(* IEC 61131-3 sources: volt/packages/volt-lsp-iec/test-corpus/awa-palletizer/Device/Plc Logic/Application/Library Manager/L_IE1P_ApplicationErrorsTypes, 22 files *)

(* ---- L_IE1P_ERROR.dut ---- *)
TYPE L_IE1P_ERROR :
(
	NOERROR := 0,
	MODULOAXISISREQUIRED := 17000,
	STARTPOSOUTOFCYCLELENGTH := 17003,
	CYCLELENGHTSHAVETOBEEQUAL := 17004,
	INVALIDDIRECTION := 17005,
	MARKSTACKLIMITREACHED := 17006,
	MAXMISSEDMARKS := 17007,
	INVALIDFOLLOWLINEACCVEL := 17008,
	INVALIDJOGGINGACCVEL := 17009,
	INVALIDSTOPDEC := 17010,
	INVALIDDIAMETER := 17011,
	TORQUEFOLLOWERNOTREADYFORMOTION := 17012,
	SPEEDFOLLOWERNOTREADYFORMOTION := 17013,
	INVALIDINVERTER := 17014,
	SDO_ACCESSFAILEDTOMOTORPARAMETERS := 17015,
	MISSEDMAPPINGPARAMETERLOWERSPEEDLIMIT := 17016,
	MISSEDMAPPINGPARAMETERUPPERSPEEDLIMIT := 17017,
	MISSEDMAPPINGPARAMETERTORQUEOFFSET := 17018,
	DANCERPOSOUTOFRANGE := 17019,
	INVALIDLIMITDANCERPOS := 17020,
	INVALIDCLUTCHPARAMETERS := 17021,
	WASNOTCALLEDDURINGMOTION := 17022,
	INVALIDNUMBEROFCAMPOINTS := 17030,
	INVALIDPATHPAR := 17032,
	INVALIDBLENDINGRADIUS := 17033,
	PATHNOTSUPPORTED := 17034,
	X_PATHLIMITPOSITIVEEXCEEDED := 17035,
	X_PATHLIMITNEGATIVEEXCEEDED := 17036,
	Y_PATHLIMITPOSITIVEEXCEEDED := 17037,
	Y_PATHLIMITNEGATIVEEXCEEDED := 17038,
	Z_PATHLIMITPOSITIVEEXCEEDED := 17039,
	Z_PATHLIMITNEGATIVEEXCEEDED := 17040,
	C_PATHLIMITPOSITIVEEXCEEDED := 17041,
	C_PATHLIMITNEGATIVEEXCEEDED := 17042,
	INVALIDPATHDATA := 17043,
	INVALIDTARGETPLC := 17047,
	MINLIMITVELGTPROFILEVEL := 17048,
	MINLIMITACCGTPROFILEACC := 17049,
	MINLIMITDECGTPROFILEDEC := 17050,
	MASTERISMOVING := 17100,
	INVALIDPODUCTLENGTH := 17101,
	TPSENSORNOTTEACHED := 17102,
	SLAVERECEIVEDGAPS := 17103,
	MASTERRECEIVEDGAPS := 17104,
	INTERNALERROR := 17105,
	INVALIDPARAMETERCUTTINGANGLE := 17106,
	INVALIDCUTTINGPARAMETERS := 17107,
	INVALIDCUTTINGLENGTH := 17108,
	SLAVENOTINPARKPOS := 17109,
	MASTERISREVERSING := 17110,
	INTINVALIDSELECTCAM := 17111,
	SELECTEDAXISISNOTSUPPORTED := 17112,
	AXISISNOTSUPPORTED := 17113,
	INVALIDPROFILE := 17114,
	AXISENABLEDISREQUIRED := 17115,
	CORRLIMITOUTOFCYCLELENGTH := 17116,
	CORRECTIONGREATERCORRWINDOW := 17117,
	INVALIDCNCPROGRAM := 17118,
	SAFEDISTVIOLATION := 17119,
	SAFEDISTINSUFFICIENTFORSTOP := 17120,
	INVALIDGCODELINE := 17121,
	COORDSYSTEMACSNOTSUPPORTED := 17122,
	DANCERLIMITSNOTTEACHED := 17123,
	NOTREADYFORADDPROFILE := 17124,
	SLAVEPOSUPPERLIMIT := 17125,
	SLAVEPOSLOWERLIMIT := 17126,
	TARGETPOSUPPERLIMIT := 17127,
	INVALIDMARKPOSITION := 17128,
	INVALIDPOSITIONINGMODE := 17129,
	TEMPSENSORFAILURE := 17130,
	MAXCRITICALTEMPREACHED := 17131,
	INVALIDTEMPCONTROLPARAM := 17132,
	IDENTIFICATIONFAILED := 17133,
	PWMTASKCYCLEMISMATCH := 17134,
	CONCURRENTREQUESTTEMPCONTROL := 17135,
	TMNOTCALLEDINCYCLICTASK := 17136,
	TMDATABUSDISCONNECTED := 17137,
	INVALIDTMDATABUS := 17138,
	TMDATABUSCONFIGCHANGED := 17139,
	TMNOTCALLEDINMOTIONTASK := 17140,
	SLAVETMSTATESERVICE := 17141,
	COLLISIONDETECTIONDISABLED := 17142,
	COLLISIONDETECTED := 17143,
	INVALIDTMDATABUSORDER := 17144,
	CHANGEOFCONVEYORAXESNOTALLOWED := 17145,
	INVALIDSETTARGET := 17146,
	LOWERLIMITEXCEEDSUPPERLIMIT := 17147,
	SETTARGETSTACKLIMITREACHED := 17148,
	WORKPIECESTACKLIMITREACHED := 17149,
	INVALIDTRAVERSINGPROFILEPARAMETER := 17150,
	INVALIDTRAVERSINGCOILPARAMETER := 17151,
	TRAVERSINGANGULARSHIFTLIMITREACHED := 17152,
	AXESGROUPALREADYINUSE := 17153,
	UNDERVOLTAGEDCLINK := 17154,
	COUPLINGMODEREQUIRESMODULOAXIS := 17155,
	DUPLICATEDTM_ADDRESS := 17156,
	XAXISTMERROR := 17157,
	YAXISTMERROR := 17158,
	APAXISTMERROR := 17159,
	SLAVEXAXISTMERROR := 17160,
	SLAVEYAXISTMERROR := 17161,
	INVALIDMOVEPPACTIVE := 17162,
	INVALIDCONVEYORBELTPAR := 17163,
	IDENTIFICATIONDIAMETERFAILED := 17164,
	ACTDANCERPOSGTMAXDANCERPOS := 17165,
	INVALIDIDENTMAXDANCERPOS := 17166,
	INVALIDDANCERMATERIALLENGTH := 17167,
	LOADDIAMETERNOTALLOWED := 17168,
	INVALIDMASTERAXISREF := 17169,
	SYNCMODEVELACCREQUIRED := 17170,
	TEMPMAXCRITICALEXCEEDED := 17171,
	INVALIDTEMPCTRLPARAM := 17172,
	INVALIDSYNCSLAVEDIRECTION := 17173,
	MARKCORRECTIONINNEXTCYCLE := 17174,
	BASEVELOCITYNOTSUPPORTED := 17175,
	MOVEMENTBLOCKEDBYTRAINAHEAD := 17176,
	MARKDISTANCEGTZEROREQUIRED := 17177,
	INVALIDVIRTMASTERSETVELZERO := 17178,
	HOMINGBLOCKEDBYACTIVEFUNCTION := 17179,
	CONCURRENTMOTIONCMDDURINGHOMING := 17180,
	INVALIDCYCLELENGTHETCONBOARD := 17181,
	INVALIDMASTERVALUESOURCE := 17182,
	ETCONBOARDNOTOPERATIONAL := 17183,
	TRAVERSINGRANGEMASTERNOTEQUALVIRTMASTER := 17184,
	CYCLELENGTHMASTERNOTEQUALVIRTMASTER := 17185,
	MISSEDMAPPINGPARAMETERTPTIMESTAMP := 17186,
	TOLERANCEALLOWEDDIRECTIONEXCEEDED := 17187,
	TPRECPOSITIONNOTSUPPORTED := 17188,
	INVALIDHYSTERESISWIDTH := 17189,
	ALLOWEDDIRECTIONVIOLATEDBYBASEVELOCITY := 17190,
	VELOUTOFTOLERANCEINVERTGEARFACTOR := 17191,
	INVALIDPARAMETERCOMBINATIONACDRIVEPROFILE := 17192,
	MINVELLIMITGTMAXVELLIMIT := 17193,
	SETVALUEMODENOTSUPPORTED := 17194,
	LINEVELDIAMCALCREQUIRED := 17195,
	INVALIDSTOPMODE := 17196,
	INVALIDDIRECTIONFORTARGETMATERIALCOUNTER := 17197,
	MAXMISSEDMARKSTOOL := 17198,
	MODECHANGEBLOCKEDBYSYNCIN := 17199,
	CONCURRENTMOTIONCMDDURINGSERVICE := 17200,
	STOPPOSITIONEXCEEDED := 17201,
	NOTREADYFORCOORDINATEDMOTION := 17202,
	INVALIDMARKWINDOWMASTERVALUECORR := 17203,
	INVALIDMARKWINDOWTOOLCORR := 17204,
	FUNCTIONBLOCKEDBYTRAVERSING := 17205,
	MASTERCYCLELENGTHCHANGED := 17206,
	TRIMMINGONLYDURINGSYNCHRONISED := 17207,
	LOWERTURNPOSGTUPPERTURNPOS := 17208,
	MASTERNOTCONNECTED := 17209,
	CANNOTCATCHUP := 17210,
	MISSINGMMADDRESS := 17901,
	NUMOFMMEXCEEDED := 17902,
	DUPLICATEDROOTMM := 17903,
	SLAVEMMNOTFOUND := 17904,
	ZPOSMAXEXCEEDED := 17905,
	MISSINGMODULEREFERENCE := 17906,
	ERRORLISTOVERFLOW := 17907,
	ACDOWNSTRUCTINVALID := 17908,
	ACDSLAVESTRUCTINVALID := 17909,
	ACDSIZEOVERFLOW := 17910,
	COMPIDOUTOFRANGE := 17911,
	TOOMANYLEVELS := 17912,
	MMDSTRUCTINVALID := 17913,
	NOPOOLRESOURCEAVAILABLE := 17914,
	NORESOURCEMOVELINABS := 17915,
	NORESOURCEMOVELINREL := 17916,
	NORESOURCEMOVEDIRABS := 17917,
	NORESOURCEMOVEDIRREL := 17918,
	NORESOURCEPNP := 17919,
	NOCOMMANDRECEIVERAVAILABLE := 17920,
	COMMANDRECEIVERNOTENABLED := 17921,
	INTERNALCONTROLACTIVE := 17922,
	INTERNALCONTROLENABLED := 17923,
	INTERNALCONTROLDISABLED := 17924,
	MMCOUPLINGDISABLED := 17925,
	MMCOUPLINGENABLED := 17926,
	MODECHANGEREQUESTED := 17927,
	MODENUMBEROUTSIDERANGE := 18001,
	MODENUMBERNOTUSEDINCONFIG := 18002,
	MODECHANGENOTALLOWEDINCURRENTMODE := 18003,
	MODECHANGENOTALLOWEDINNEXTMODE := 18004,
	LI_MODENUMBEROUTSIDERANGE := 18005,
	LI_MODENUMBERNOTUSEDINCONFIG := 18006,
	LI_MODECHANGENOTALLOWEDREMOTE := 18007,
	LI_MODECHANGENOTALLOWEDINCURRENTMODE := 18008,
	LI_MODECHANGENOTALLOWEDINNEXTMODE := 18009,
	MORETHANONECOMMANDACTIVE := 18010,
	CONCURRENTCOMMAND := 18011,
	COMMANDNOTALLOWEDINCURRENTSTATE := 18012,
	LI_COMMANDSONLYINMODEPRODUCTION := 18013,
	LI_COMMANDNOTALLOWEDINREMOTE := 18014,
	LI_COMMANDNOTALLOWEDINCURRENTSTATE := 18015,
	CONCURRENTTOOLCMD := 18016,
	DELAYTIMEINVALID_PT1FILTER := 19000,
	MODEINVALID_CURVE := 19002,
	MODEINVALID_COMPARE := 19003,
	MODEINVALID_CONVAXISV := 19005,
	DELAYTIMEINVALID_PROCESSCONTROLLER := 19006,
	RATETIMEINVALID_PROCESSCONTROLLER := 19007,
	RESETTIMEINVALID_PROCESSCONTROLLER := 19008,
	MODEINVALID_DELAY := 19024,
	ABORTEDBYSTARTIDENT_FRICTCOMP := 19030,
	ABORTEDBYFOLLOWERDISABLED_FRICTCOMP := 19031,
	MAXSPEEDNOTREACHED_FRICTCOMP := 19032,
	ACCTOOBIG_FRICTCOMP := 19033,
	DMINBIGGERDMAX_CALCDIAMETER := 19034,
	MAXSPEEDORMAXTORQUE_IDENTMINERTIA := 19048,
	ABORTEDBYSTARTIDENT_IDENTMINERTIA := 19049,
	ABORTEDBYFOLLOWERDISABLED_IDENTMINERTIA := 19050,
	ABORTEDBYFOLLOWERENABLED_IDENTMINERTIA := 19051,
	NMAXNOTREACHED_IDENTMINERTIA := 19052,
	MNOTREACHED_IDENTMINERTIA := 19053,
	MAXNROFTPEXCEEDED_MARKREGISTER := 19503,
	IDENTMODENOTSUPPORTED := 19801,
	MOTORRATEDSPEEDZERO := 19803,
	INERTIAMOTORZERO := 19804,
	STARTMODEINVALID := 19806,
	INVALIDEIGENFREQUENCY := 19807,
	INVALIDAMPLITUDERATIO := 19808,
	INVALIDOSCCOMPMODE := 19809,
	CHANGEOFOSCCOMPMODELOCKED := 19810,
	INVALIDDEFAULTCONTROLMODE := 19812,
	INVALIDMOTORCONTROLMODE := 19813,
	VIRTUALMODENOTALLOWED := 19814,
	POSITIONWINDOWNEGOUTSIDESWLIMITS := 19817,
	POSITIONWINDOWPOSOUTSIDESWLIMITS := 19818,
	ACTPOSITIONOUTSIDEWINDOW := 19819,
	PROFILEEXCEEDSPOSITIONWINDOW := 19820,
	ACTVELOCITYEXCEEDSTOLERANCE := 19822,
	ACTTORQUEEXCEEDSTOLERANCE := 19823,
	POSITIONWINDOWNEGVIOLATION := 19825,
	POSITIONWINDOWPOSVIOLATION := 19826,
	AXISINSTABILITYDUETOSTARTCTRLPARAM := 19827,
	INPOSITIONTIMEOUT := 19828,
	RESTOREDATANOTAVAILABLE := 19829,
	POSITIONWINDOWREQUIRESLIMITEDAXIS := 19830,
	MISSEDMAPPINGPARAMETERVELOCITYERROR := 19831,
	INSTABILITYDUETOTUNESTRATEGY := 19832,
	ARRAYBOUNDSNOTEQUALMODULOCYCLE := 19833,
	PERIODICCORRECTIONVALUESREQUIRED := 19834,
	INVALIDBACKLASHCOMPMODE := 19835,
	INVALIDBACKLASHWIDTH := 19836,
	INVALIDCOMPTIME := 19837,
	BACKLASHWIDTHGTCYCLELENGTH := 19838,
	SDO_OTHERERROR := 20001,
	SDO_INVALIDINDEX := 20002,
	SDO_INVALIDOFFSET := 20003,
	SDO_INVALIDSIZE := 20004,
	SDO_INVALIDDATA := 20005,
	SDO_NOTREADY := 20006,
	SDO_BUSY := 20007,
	SDO_NOMEMORY := 20008,
	SDO_INVALIDPARM := 20009,
	SDO_INVALIDSTATE := 20010,
	SDO_TIMEOUT := 20011,
	SDO_INVALID_SLAVE_STATE := 20012,
	SDO_LINK_DISCONNECTED := 20013,
	SDO_ALL_CANNELS_BUSY := 20015,
	SDO_ABORTCODE_TOGGLE := 20020,
	SDO_ABORTCODE_TIMEOUT := 20021,
	SDO_ABORTCODE_CCS_SCS := 20022,
	SDO_ABORTCODE_BLK_SIZE := 20023,
	SDO_ABORTCODE_SEQNO := 20024,
	SDO_ABORTCODE_CRC := 20025,
	SDO_ABORTCODE_MEMORY := 20026,
	SDO_ABORTCODE_ACCESS := 20027,
	SDO_ABORTCODE_WRITEONLY := 20028,
	SDO_ABORTCODE_READONLY := 20029,
	SDO_ABORTCODE_INDEX := 20030,
	SDO_ABORTCODE_PDO_MAP := 20031,
	SDO_ABORTCODE_PDO_LEN := 20032,
	SDO_ABORTCODE_P_INCOMP := 20033,
	SDO_ABORTCODE_I_INCOMP := 20034,
	SDO_ABORTCODE_HARDWARE := 20035,
	SDO_ABORTCODE_DATA_SIZE := 20036,
	SDO_ABORTCODE_DATA_SIZE1 := 20037,
	SDO_ABORTCODE_DATA_SIZE2 := 20038,
	SDO_ABORTCODE_OFFSET := 20039,
	SDO_ABORTCODE_DATA_RANGE := 20040,
	SDO_ABORTCODE_DATA_RANGE1 := 20041,
	SDO_ABORTCODE_DATA_RANGE2 := 20042,
	SDO_ABORTCODE_MINMAX := 20043,
	SDO_ABORTCODE_GENERAL := 20044,
	SDO_ABORTCODE_TRANSFER := 20045,
	SDO_ABORTCODE_TRANSFER1 := 20046,
	SDO_ABORTCODE_TRANSFER2 := 20047,
	SDO_ABORTCODE_DICTIONARY := 20048,
	SDO_ABORTCODE_UNKNOWN := 20049,
	NOAXISREF := 20301,
	NOPARAMETER := 20302,
	NOVALIDPARAM := 20303,
	NOVALIDAXISSTATE := 20304,
	NOBOOLPARAM := 20305,
	SWLIMITPOS := 20306,
	SWLIMITNEG := 20307,
	NOVALID_MC_SOURCE := 20308,
	NOSETVALUESAVAILABLE := 20309,
	POWERFAILDURINGOPERATION := 20310,
	NOTREADYFORMOTION := 20311,
	POSSWLIMITREACHED := 20312,
	NEGSWLIMITREACHED := 20313,
	NOVALIDTPSOURCE := 20314,
	NOVALIDTPNUMBER := 20315,
	TPALREADYACTIVE := 20316,
	NOTTPSUPPORTED := 20317,
	NOTPACTIVE := 20318,
	NOEXTPINPUT := 20319,
	NOVALIDACCELERATION := 20320,
	NOVALIDDECELERATION := 20321,
	NOVALIDVELOCITY := 20322,
	ARITHMETICERROR := 20323,
	NOTAPPLICABLE := 20324,
	VELOCITYLIMITED := 20325,
	ACCELERATIONLIMITED := 20326,
	JERKLIMITED := 20327,
	TARGETOUTSIDESWLIMIT := 20328,
	JERKLIMITATIONDEACTIVATEDDUETOARITHMETICERROR := 20329,
	NOVALIDACCELERATION_MOVEABSOLUTE := 20330,
	NOVALIDDECELERATION_MOVEABSOLUTE := 20331,
	NOVALIDVELOCITY_MOVEABSOLUTE := 20332,
	ARITHMETICERROR_MOVEABSOLUTE := 20333,
	NOTAPPLICABLE_MOVEABSOLUTE := 20334,
	VELOCITYLIMITED_MOVEABSOLUTE := 20335,
	ACCELERATIONLIMITED_MOVEABSOLUTE := 20336,
	JERKLIMITED_MOVEABSOLUTE := 20337,
	TARGETOUTSIDESWLIMIT_MOVEABSOLUTE := 20338,
	NOVALIDACCELERATION_MOVEADDITIVE := 20340,
	NOVALIDDECELERATION_MOVEADDITIVE := 20341,
	NOVALIDVELOCITY_MOVEADDITIVE := 20342,
	ARITHMETICERROR_MOVEADDITIVE := 20343,
	NOTAPPLICABLE_MOVEADDITIVE := 20344,
	VELOCITYLIMITED_MOVEADDITIVE := 20345,
	ACCELERATIONLIMITED_MOVEADDITIVE := 20346,
	JERKLIMITED_MOVEADDITIVE := 20347,
	TARGETOUTSIDESWLIMIT_MOVEADDITIVE := 20348,
	NOVALIDACCELERATION_MOVECONTAB := 20350,
	NOVALIDDECELERATION_MOVECONTAB := 20351,
	NOVALIDVELOCITY_MOVECONTAB := 20352,
	ARITHMETICERROR_MOVECONTAB := 20353,
	NOTAPPLICABLE_MOVECONTAB := 20354,
	VELOCITYLIMITED_MOVECONTAB := 20355,
	ACCELERATIONLIMITED_MOVECONTAB := 20356,
	JERKLIMITED_MOVECONTAB := 20357,
	TARGETOUTSIDESWLIMIT_MOVECONTAB := 20358,
	NOVALIDACCELERATION_MOVECONTREL := 20360,
	NOVALIDDECELERATION_MOVECONTREL := 20361,
	NOVALIDVELOCITY_MOVECONTREL := 20362,
	ARITHMETICERROR_MOVECONTREL := 20363,
	NOTAPPLICABLE_MOVECONTREL := 20364,
	VELOCITYLIMITED_MOVECONTREL := 20365,
	ACCELERATIONLIMITED_MOVECONTREL := 20366,
	JERKLIMITED_MOVECONTREL := 20367,
	TARGETOUTSIDESWLIMIT_MOVECONTREL := 20368,
	NOVALIDACCELERATION_MOVERELATIVE := 20370,
	NOVALIDDECELERATION_MOVERELATIVE := 20371,
	NOVALIDVELOCITY_MOVERELATIVE := 20372,
	ARITHMETICERROR_MOVERELATIVE := 20373,
	NOTAPPLICABLE_MOVERELATIVE := 20374,
	VELOCITYLIMITED_MOVERELATIVE := 20375,
	ACCELERATIONLIMITED_MOVERELATIVE := 20376,
	JERKLIMITED_MOVERELATIVE := 20377,
	TARGETOUTSIDESWLIMIT_MOVERELATIVE := 20378,
	NOVALIDACCELERATION_MOVESUPERIMP := 20380,
	NOVALIDDECELERATION_MOVESUPERIMP := 20381,
	NOVALIDVELOCITY_MOVESUPERIMP := 20382,
	ARITHMETICERROR_MOVESUPERIMP := 20383,
	NOTAPPLICABLE_MOVESUPERIMP := 20384,
	VELOCITYLIMITED_MOVESUPERIMP := 20385,
	ACCELERATIONLIMITED_MOVESUPERIMP := 20386,
	JERKLIMITED_MOVESUPERIMP := 20387,
	TARGETOUTSIDESWLIMIT_MOVESUPERIMP := 20388,
	NOVALIDACCELERATION_MOVEVELOCITY := 20390,
	NOVALIDDECELERATION_MOVEVELOCITY := 20391,
	NOVALIDVELOCITY_MOVEVELOCITY := 20392,
	ARITHMETICERROR_MOVEVELOCITY := 20393,
	NOTAPPLICABLE_MOVEVELOCITY := 20394,
	VELOCITYLIMITED_MOVEVELOCITY := 20395,
	ACCELERATIONLIMITED_MOVEVELOCITY := 20396,
	JERKLIMITED_MOVEVELOCITY := 20397,
	TARGETOUTSIDESWLIMIT_MOVEVELOCITY := 20398,
	NOVALIDDECELERATION_HALT := 20401,
	ARITHMETICERROR_HALT := 20403,
	ACCELERATIONLIMITED_HALT := 20406,
	JERKLIMITED_HALT := 20407,
	NOVALIDDECELERATION_STOP := 20411,
	ARITHMETICERROR_STOP := 20413,
	ACCELERATIONLIMITED_STOP := 20416,
	JERKLIMITED_STOP := 20417,
	NOVALIDDIRECTION := 20430,
	NOVALIDBUFFERMODE := 20431,
	DIRECTIONDISABLED := 20432,
	BLOCKEDBYAXISSTATE := 20433,
	NOVALIDOVERRIDE := 20434,
	CONCURRENT_MC_POWER := 20435,
	CONCURRENT_SETQUICKSTOP := 20436,
	FDBABSPOSNOTAVAILABLE := 20498,
	DRIVE_PDO_INTERFACE_DISABLED := 20499,
	HWLIMITPOS := 20500,
	HWLIMITNEG := 20501,
	FOLLOWINGERROR1 := 20502,
	FOLLOWINGERROR2 := 20503,
	COMMUNICATIONFAIL := 20504,
	AXISINITFAIL := 20505,
	COMMTIMOUT := 20506,
	MASTERRESTARTFAIL := 20507,
	NOTREADYFORREINIT := 20508,
	ERRORDURINGINIT := 20509,
	SWITCHONNOTPOSSIBLE := 20510,
	DRIVEERROR := 20511,
	HOME_NOAUXPARAMETERS := 20512,
	HOME_MODENOTSUPPORTEDBYAXIS := 20513,
	HOME_MODEUNKNOWN := 20514,
	HOME_NOAUXTRIGGERINPUT := 20515,
	HOME_UNKNOWNTPCONFIG := 20516,
	HOME_WRITEHOMEPARAMETER := 20518,
	HOME_ERRORWHILEHOMING := 20519,
	HOME_ARITHMETICERROR := 20520,
	HOME_TORQUELIMNOTMAPPED := 20521,
	HOME_INVALIDVELACC := 20522,
	HOMETPEDGESETTINGNOTSUPPORTED := 20523,
	RESETDRIVEERRORFAILED := 20525,
	APPLICATIONERROR := 20526,
	APPLICATIONWARNING := 20527,
	BRAKE_POSITIONDRIFT := 20529,
	BRAKE_INVALIDMODE := 20530,
	BRAKE_TIMEOUTPRECONTROL := 20531,
	BRAKE_INVALIDBRAKESTATE := 20532,
	FAST_IO_OUT_WRONGOUTPUTSEL := 20533,
	FAST_IO_OUT_NOFREEENCODERAXIS := 20534,
	FAST_IO_OUT_FREEENCODERAXISWRONGPARAMETER := 20535,
	FAST_IO_OUT_MAPPINGFAULT := 20536,
	FAST_IO_OUT_FIFOOVERFLOW := 20537,
	TP_SELECT := 20538,
	TP_MODE := 20539,
	TP_ONLYPOSEDGE := 20540,
	TP_EDGENOTAVAILABLE := 20541,
	TP_CHANNELNOTFREE := 20542,
	TP_MAPPINGFAULT := 20543,
	TP_INTERNALCHANNELNOTFREE := 20544,
	TP_TIMEOUT := 20545,
	TP_COMMUNICATIONERROR := 20546,
	TP_SIGNAL := 20547,
	TP_NOFREEENCODERAXIS := 20548,
	TP_PARAMETERRISINGEDGEWRONGVALUE := 20550,
	TP_PARAMETERFALLINGRISINGEDGEWRONGVALUE := 20551,
	TP_INTERNALERROR := 20552,
	SETVALUESGTMAXAPPVALUES := 20600,
	SETVALUESINCONSISTENT := 20601,
	POSDIFFGTHALFCYCLELENGTH := 20602,
	INVALIDTASKCYCLETIME := 20603,
	INIT_WRITEERRORSDO := 20650,
	INIT_READERRORSDO := 20651,
	INIT_MAXTASKTIME := 20652,
	INIT_TORQUEREFISZERO := 20653,
	INIT_MOTORRATEDSPEEDISZERO := 20654,
	INIT_REVISIONNOTVALID := 20655,
	INIT_ENCCOUNTNOTVALID := 20656,
	INIT_ENCREVNOTVALID := 20657,
	INIT_ENCCRCNOTVALID := 20658,
	INIT_ENCABSPOSNOTAVAILABLE := 20659,
	CONTROLLERFIRMWARENOTCOMPATIBLE := 20660,
	INVALIDMODE := 20661,
	ENCBPB_INIT_FAILED := 20662,
	LEDNOTSUPPORTEDBYDEVICE := 20663,
	INVALIDGEARFACTOR := 20664,
	POSOUTOFCYCLELENGTH := 20665,
	CYCLELENGTHINVALID_ADDOFFSETCYCLIC := 20666,
	POSININVALID_ADDOFFSETCYCLIC := 20667,
	CYCLELENGTHINVALID_ZERODETECT := 20668,
	POSININVALID_ZERODETECT := 20669,
	STARTPOSINVALID_INTEGRATEAXIS := 20670,
	INVALIDINPUTJOGPOSJOGNEG := 20671,
	VALUEOUTOFRANGE := 20672,
	STATENOTEQUALDISABLED := 20673,
	INVALIDINPUT_BRAKETEST := 20674,
	ALREADYACTIVE_BRAKETEST := 20675,
	INVALIDINPUT_BRAKEGRINDIN := 20676,
	ALREADYACTIVE_GRINDIN := 20677,
	INVALIDCONTROLMODE := 20678,
	VIRTUALAXISNOTSUPPORTED := 20679,
	AXISNOTDISABLED := 20680,
	INVALIDFEEDCONSTANT := 20681,
	INVALIDTRAVERSINGRANGE := 20682,
	INVALIDCYCLELENGTH := 20683,
	INVALIDPOSRESOLUTION := 20684,
	TORQUELIMTOOLARGE := 20685,
	TORQUELIMLESSTHANZERO := 20686,
	INVALIDLOADENCSIGNAL := 20687,
	ENCSIGNALGTMEASURINGRANGE := 20688,
	INVALIDENCMEASURINGRANGE := 20689,
	DRIVESTOACTIVE := 20690,
	DRIVECINHACTIVE := 20691,
	INVALIDSWLIMITS := 20692,
	NOVALIDJERK := 20693,
	MISSEDMAPPINGPARAMETERVLTARGETVEL := 20694,
	MISSEDMAPPINGPARAMETERVLACTUALVEL := 20695,
	AXISNOTHOMED := 20696,
	AXISNOTINSIMPLEMODE := 20697,
	AXISINSIMPLEMODE := 20698,
	FUNCTIONNOTSUPPORTEDBYAXIS := 20699,
	EXECUTIONINDEXALREADYINUSE := 20700,
	SS1ACTIVE := 20701,
	SS2ACTIVE := 20702,
	VELOCITYLIMITEDBYSLS1 := 20703,
	VELOCITYLIMITEDBYSLS2 := 20704,
	VELOCITYLIMITEDBYSLS3 := 20705,
	VELOCITYLIMITEDBYSLS4 := 20706,
	INVALIDEXECUTIONINDEX := 20707,
	INVALIDFILTERDEPTH := 20708,
	PARAMSETFAILEDJOGVEL := 20709,
	PARAMSETFAILEDJOGACC := 20710,
	PARAMSETFAILEDJOGDEC := 20711,
	PARAMSETFAILEDJOGJERK := 20712,
	PARAMSETFAILEDHALTDEC := 20713,
	PARAMSETFAILEDHALTJERK := 20714,
	PARAMSETFAILEDQSPAPPLDEC := 20715,
	PARAMSETFAILEDQSPAPPLJERK := 20716,
	PARAMSETFAILEDHOMEPOSITION := 20717,
	PARAMSETFAILEDHOMEMODE := 20718,
	PARAMSETFAILEDHOMESTOPMODE := 20719,
	PARAMSETFAILEDHOMETARGETPOSITION := 20720,
	PARAMSETFAILEDHOMEVELOCITY1 := 20721,
	PARAMSETFAILEDHOMEVELOCITY2 := 20722,
	PARAMSETFAILEDHOMEACCELERATION1 := 20723,
	PARAMSETFAILEDHOMEACCELERATION2 := 20724,
	PARAMSETFAILEDHOMEJERK := 20725,
	PARAMSETFAILEDHOMETORQUELIMIT := 20726,
	PARAMSETFAILEDHOMETORQUETIME := 20727,
	PARAMSETFAILEDHOMETPCONFIG := 20728,
	PARAMSETFAILEDDRIVEHOMEMODE := 20729,
	PARAMREADFAILED := 20730,
	PARAMROLLBACKFAILED := 20731,
	POSCTRLNOTSUPPORTED := 20732,
	TORQUECTRLNOTSUPPORTED := 20733,
	SETPOSITIONINPDOREQUIRED := 20734,
	SETVELOCITYINPDOREQUIRED := 20735,
	SETTORQUEINPDOREQUIRED := 20736,
	UPPERSPEEDLIMINPDOREQUIRED := 20737,
	LOWERSPEEDLIMINPDOREQUIRED := 20738,
	ACTPOSITIONINPDOREQUIRED := 20739,
	BRAKEGRINDININVALIDPOSITIONLIMITS := 20740,
	BRAKEGRINDINSTARTPOSOUTSIDEPOSLIM := 20741,
	BRAKEGRINDINDISTANCENOTSUFFICIENT := 20742,
	SAFETYNOTSUPPORTEDBYDRIVE := 20743,
	SAFETYCONTROLWORDINPDOREQUIRED := 20744,
	SETPOSITIONONSLAVEAXISNOTALLOWED := 20745,
	ENCODERVELOCITYGTMAXVELOCITY := 20746,
	INVALIDENCODERSIGNAL := 20747,
	DRIVESAFEBRAKECTRLACTIVE := 20748,
	POSRECONSTRMAXAXISREACHED := 20749,
	POSRECONSTRDATAINKONSISTENT := 20750,
	POSRECONSTRHOMEPOSAVAILABLENOTACTIVE := 20751,
	POSRECONSTRNOTACTIVATED := 20752,
	POSRECONSTRAXISWASVIRTUAL := 20753,
	POSRECONSTRORIENTATIONCHANGED := 20754,
	POSRECONSTRTRAVERSINGRANGECHANGED := 20755,
	POSRECONSTRCYCLELENGTHCHANGED := 20756,
	POSRECONSTRUNITFACTORCHANGED := 20757,
	POSRECONSTRRESETBYENCERROR := 20758,
	POSRECONSTRRESETBYFDBCHANGED := 20759,
	POSRECONSTRENCCRCCHANGED := 20760,
	POSRECONSTRNOFDBPOSAVAILABLE := 20761,
	POSRECONSTRABSENCREQUIRED := 20762,
	POSRECONSTRDATAVERSIONCHANGED := 20763,
	POSRECONSTRNODATAAVAILABLE := 20764,
	POSRECONSTRNOMEMORYAVAILABLE := 20765,
	POSRECONSTRPOSOUTSIDERESTORETRESHOLD := 20766,
	POSRECONSTRRESETBYFDBOPENCIRC := 20767,
	PPIMODENOTSUPPORTED := 20768,
	PPINOTSUCCESSFULL := 20769,
	POLEPOSITIONNOTAVAILABLE := 20770,
	CONCURRENTPPI := 20771,
	PARAMNOTACCESSIBLE := 20773,
	MISSINGMAPPINGPARAMETER := 20774,
	PARAMUSEDBYAXISREF := 20775,
	PARAMMAPPEDWITHWRITEACCESS := 20776,
	PARAMMAPPEDWITHREADACCESS := 20777,
	MOLMODENOTSUPPORTED := 20778,
	HOMEPOSRESETBYMACHINEDATACHANGEAPPL := 20779,
	HOMEPOSRESETBYMACHINEDATACHANGE := 20780,
	HOMEPOSRESETBYENCCRCCHANGED := 20781,
	HOMEPOSRESETBYDRIVESWITCHEDOFF := 20782,
	HOMEPOSRESETBYFDBCHANGED := 20783,
	HOMEPOSRESETBYFDBABSPOSNOTAVAILABLE := 20784,
	HOMEPOSRESETBYENCERROR := 20785,
	HOMEPOSRESETBYAPPLICATION := 20786,
	HOMEPOSRESETBYFDBOPENCIRC := 20787,
	HOMEPOSRESETBYSTARTREFERENCESEARCH := 20788,
	HOMEPOSRESETBYVIRTUALMODE := 20789,
	HOMEPOSRESETBYAXESGROUP := 20790,
	POSRECONSTRSUCCEDED := 20791,
	HOMEPOSSETDIRECT := 20792,
	HOMEPOSSETBYREFERENCESEARCH := 20793,
	HOMEPOSSETBYAXESGROUP := 20794,
	REFERENCESEARCHABORTED := 20795,
	AXISPERSISTENTMEMORYNOTAVAILABLE := 20796,
	AXISPERSISTENTMEMORYINVALID := 20797,
	AXISPERSISTENTMEMORYNOTINITIALIZED := 20798,
	POSRECONSTRDATANOTINITIALIZED := 20799,
	MISSEDMAPPINGPARAMETERPOSTORQUELIMIT := 20800,
	MISSEDMAPPINGPARAMETERNEGTORQUELIMIT := 20801,
	MISSEDMAPPINGPARAMETERACTUALPOS := 20802,
	AUTOTUNINGNOTSUPPORTEDBYFIRMWAREVERSION := 20803,
	AUTOTUNINGEXECUTEDVARIABLESWITCHINGFREQUENCY := 20804,
	CONCURRENTREQUESTSERVICEFUNCTION := 20805,
	SETPOSNOTALLOWEDHOMEPOSPERMANENTLYSET := 20806,
	EXTENCODERREQUIREDBYPOSCTRL := 20807,
	PARAMSETFAILEDHOMEOFFSETPOS := 20808,
	PARAMSETFAILEDHOMESTOPMODEDIR := 20809,
	TORQUENOTREACHEDBRAKETEST := 20810,
	INVALIDABSPOSEXTENC := 20811,
	EXTENCODERVELOCITYGTMAXVELOCITY := 20813,
	MAXCYCLICREADCOUNTEXCEEDED := 20814,
	MAXCYCLICWRITECOUNTEXCEEDED := 20815,
	CYCLICPARAMACCESSSTILLBUSY := 20816,
	CONCURRENTCYCLICWRITEACCESS := 20817,
	BRAKETESTSUCCESSFUL := 20818,
	SBCREQUESTED := 20820,
	JOGGINGLIMITEDBYSLI := 20821,
	BRAKEGRINDINDONE := 20822,
	BRAKEGRINDINABORTED := 20823,
	BRAKETESTABORTED := 20824,
	AUTOTUNINGDONE := 20825,
	AUTOTUNINGABORTED := 20826,
	TIMESTAMPNOTSUPPORTEDBYSOURCE := 20828,
	INVALIDTIMEDELAY := 20829,
	DRIVEERRORMSGNOTRESOLVABLE := 20830,
	DRIVEWARNINGMSGNOTRESOLVABLE := 20831,
	POSRECONSTRCONNECTEDDRIVECHANGED := 20832,
	AXESCONTROLMODENOTEQUAL := 20833,
	AXESSPEEDFILTERTIMENOTEQUAL := 20834,
	AXESMOTORNOTEQUAL := 20835,
	AXESINVERTERTANOTEQUAL := 20836,
	AXESSWITCHINGFREQNOTEQUAL := 20837,
	AXESEXTFEEDBACKCONFIGNOTEQUAL := 20839,
	SSIENCODERSTATUS1ACTIVE := 20840,
	CONNECTEDDEVICENODEDISABLED := 20841,
	ETHERCATSLAVENOTPRESENT := 20842,
	MAINAXISNOTREADY := 21001,
	GROUPSTATEUNDEFINED := 21002,
	AXISDISABLED := 21003,
	TRANSFORMATIONERROR := 21004,
	AXISINERRORSTOP := 21005,
	AXISLIMITVIOLATIONMAINAXIS := 21006,
	AXISLIMITVIOLATIONREALAXIS := 21007,
	AXISLIMITVIOLATIONPASSIVEAXIS := 21008,
	REALAXISDISABLED := 21009,
	NOVALIDPATHCOICE_MOVECIRCABS := 21010,
	NOVALIDCIRCMODE_MOVECIRCABS := 21011,
	NOVALIDTRANSITIONPARAMETER_MOVECIRCABS := 21012,
	NOVALIDVELOCITY_MOVECIRCABS := 21013,
	NOVALIDACCELERATION_MOVECIRCABS := 21014,
	NOVALIDDECELERATION_MOVECIRCABS := 21015,
	NOVALIDJERK_MOVECIRCABS := 21016,
	TARGETOUTSIDESWLIMITSPASSIVEJOINTS_MOVECIRCABS := 21017,
	TARGETOUTSIDESWLIMITSMAINAXISX_MOVECIRCABS := 21018,
	TARGETOUTSIDESWLIMITSMAINAXISY_MOVECIRCABS := 21019,
	TARGETOUTSIDESWLIMITSMAINAXISZ_MOVECIRCABS := 21020,
	TARGETOUTSIDESWLIMITSMAINAXISA_MOVECIRCABS := 21021,
	TARGETOUTSIDESWLIMITSMAINAXISB_MOVECIRCABS := 21022,
	TARGETOUTSIDESWLIMITSMAINAXISC_MOVECIRCABS := 21023,
	TARGETOUTSIDESWLIMITSREALAXIS1_MOVECIRCABS := 21024,
	TARGETOUTSIDESWLIMITSREALAXIS2_MOVECIRCABS := 21025,
	TARGETOUTSIDESWLIMITSREALAXIS3_MOVECIRCABS := 21026,
	TARGETOUTSIDESWLIMITSREALAXIS4_MOVECIRCABS := 21027,
	TARGETOUTSIDESWLIMITSREALAXIS5_MOVECIRCABS := 21028,
	TARGETOUTSIDESWLIMITSREALAXIS6_MOVECIRCABS := 21029,
	TARGETOUTSIDESWLIMITSAUXAXIS1_MOVECIRCABS := 21030,
	TARGETOUTSIDESWLIMITSAUXAXIS2_MOVECIRCABS := 21031,
	TARGETOUTSIDESWLIMITSAUXAXIS3_MOVECIRCABS := 21032,
	TARGETOUTSIDESWLIMITSAUXAXIS4_MOVECIRCABS := 21033,
	TARGETOUTSIDESWLIMITSAUXAXIS5_MOVECIRCABS := 21034,
	TARGETOUTSIDESWLIMITSAUXAXIS6_MOVECIRCABS := 21035,
	TARGETTRANSFORMATIONERROR_MOVECIRCABS := 21036,
	TARGETSINGULARPOS_MOVECIRCABS := 21037,
	BORDEROUTSIDESWLIMITSPASSIVEJOINTS_MOVECIRCABS := 21038,
	BORDEROUTSIDESWLIMITSMAINAXISX_MOVECIRCABS := 21039,
	BORDEROUTSIDESWLIMITSMAINAXISY_MOVECIRCABS := 21040,
	BORDEROUTSIDESWLIMITSMAINAXISZ_MOVECIRCABS := 21041,
	BORDEROUTSIDESWLIMITSMAINAXISA_MOVECIRCABS := 21042,
	BORDEROUTSIDESWLIMITSMAINAXISB_MOVECIRCABS := 21043,
	BORDEROUTSIDESWLIMITSMAINAXISC_MOVECIRCABS := 21044,
	BORDEROUTSIDESWLIMITSREALAXIS1_MOVECIRCABS := 21045,
	BORDEROUTSIDESWLIMITSREALAXIS2_MOVECIRCABS := 21046,
	BORDEROUTSIDESWLIMITSREALAXIS3_MOVECIRCABS := 21047,
	BORDEROUTSIDESWLIMITSREALAXIS4_MOVECIRCABS := 21048,
	BORDEROUTSIDESWLIMITSREALAXIS5_MOVECIRCABS := 21049,
	BORDEROUTSIDESWLIMITSREALAXIS6_MOVECIRCABS := 21050,
	BORDEROUTSIDESWLIMITSAUXAXIS1_MOVECIRCABS := 21051,
	BORDEROUTSIDESWLIMITSAUXAXIS2_MOVECIRCABS := 21052,
	BORDEROUTSIDESWLIMITSAUXAXIS3_MOVECIRCABS := 21053,
	BORDEROUTSIDESWLIMITSAUXAXIS4_MOVECIRCABS := 21054,
	BORDEROUTSIDESWLIMITSAUXAXIS5_MOVECIRCABS := 21055,
	BORDEROUTSIDESWLIMITSAUXAXIS6_MOVECIRCABS := 21056,
	BORDERTRANSFORMATIONERROR_MOVECIRCABS := 21057,
	BORDERSINGULARPOS_MOVECIRCABS := 21058,
	ILLEGALPARAMETER_MOVECIRCABS := 21059,
	NOVALIDPATHCOICE_MOVECIRCREL := 21060,
	NOVALIDCIRCMODE_MOVECIRCREL := 21061,
	NOVALIDTRANSITIONPARAMETER_MOVECIRCREL := 21062,
	NOVALIDVELOCITY_MOVECIRCREL := 21063,
	NOVALIDACCELERATION_MOVECIRCREL := 21064,
	NOVALIDDECELERATION_MOVECIRCREL := 21065,
	NOVALIDJERK_MOVECIRCREL := 21066,
	TARGETOUTSIDESWLIMITSPASSIVEJOINTS_MOVECIRCREL := 21067,
	TARGETOUTSIDESWLIMITSMAINAXISX_MOVECIRCREL := 21068,
	TARGETOUTSIDESWLIMITSMAINAXISY_MOVECIRCREL := 21069,
	TARGETOUTSIDESWLIMITSMAINAXISZ_MOVECIRCREL := 21070,
	TARGETOUTSIDESWLIMITSMAINAXISA_MOVECIRCREL := 21071,
	TARGETOUTSIDESWLIMITSMAINAXISB_MOVECIRCREL := 21072,
	TARGETOUTSIDESWLIMITSMAINAXISC_MOVECIRCREL := 21073,
	TARGETOUTSIDESWLIMITSREALAXIS1_MOVECIRCREL := 21074,
	TARGETOUTSIDESWLIMITSREALAXIS2_MOVECIRCREL := 21075,
	TARGETOUTSIDESWLIMITSREALAXIS3_MOVECIRCREL := 21076,
	TARGETOUTSIDESWLIMITSREALAXIS4_MOVECIRCREL := 21077,
	TARGETOUTSIDESWLIMITSREALAXIS5_MOVECIRCREL := 21078,
	TARGETOUTSIDESWLIMITSREALAXIS6_MOVECIRCREL := 21079,
	TARGETOUTSIDESWLIMITSAUXAXIS1_MOVECIRCREL := 21080,
	TARGETOUTSIDESWLIMITSAUXAXIS2_MOVECIRCREL := 21081,
	TARGETOUTSIDESWLIMITSAUXAXIS3_MOVECIRCREL := 21082,
	TARGETOUTSIDESWLIMITSAUXAXIS4_MOVECIRCREL := 21083,
	TARGETOUTSIDESWLIMITSAUXAXIS5_MOVECIRCREL := 21084,
	TARGETOUTSIDESWLIMITSAUXAXIS6_MOVECIRCREL := 21085,
	TARGETTRANSFORMATIONERROR_MOVECIRCREL := 21086,
	TARGETSINGULARPOS_MOVECIRCREL := 21087,
	BORDEROUTSIDESWLIMITSPASSIVEJOINTS_MOVECIRCREL := 21088,
	BORDEROUTSIDESWLIMITSMAINAXISX_MOVECIRCREL := 21089,
	BORDEROUTSIDESWLIMITSMAINAXISY_MOVECIRCREL := 21090,
	BORDEROUTSIDESWLIMITSMAINAXISZ_MOVECIRCREL := 21091,
	BORDEROUTSIDESWLIMITSMAINAXISA_MOVECIRCREL := 21092,
	BORDEROUTSIDESWLIMITSMAINAXISB_MOVECIRCREL := 21093,
	BORDEROUTSIDESWLIMITSMAINAXISC_MOVECIRCREL := 21094,
	BORDEROUTSIDESWLIMITSREALAXIS1_MOVECIRCREL := 21095,
	BORDEROUTSIDESWLIMITSREALAXIS2_MOVECIRCREL := 21096,
	BORDEROUTSIDESWLIMITSREALAXIS3_MOVECIRCREL := 21097,
	BORDEROUTSIDESWLIMITSREALAXIS4_MOVECIRCREL := 21098,
	BORDEROUTSIDESWLIMITSREALAXIS5_MOVECIRCREL := 21099,
	BORDEROUTSIDESWLIMITSREALAXIS6_MOVECIRCREL := 21100,
	BORDEROUTSIDESWLIMITSAUXAXIS1_MOVECIRCREL := 21101,
	BORDEROUTSIDESWLIMITSAUXAXIS2_MOVECIRCREL := 21102,
	BORDEROUTSIDESWLIMITSAUXAXIS3_MOVECIRCREL := 21103,
	BORDEROUTSIDESWLIMITSAUXAXIS4_MOVECIRCREL := 21104,
	BORDEROUTSIDESWLIMITSAUXAXIS5_MOVECIRCREL := 21105,
	BORDEROUTSIDESWLIMITSAUXAXIS6_MOVECIRCREL := 21106,
	BORDERTRANSFORMATIONERROR_MOVECIRCREL := 21107,
	BORDERSINGULARPOS_MOVECIRCREL := 21108,
	ILLEGALPARAMETER_MOVECIRCREL := 21109,
	NOVALIDTRANSITIONPARAMETER_MOVELINABS := 21110,
	NOVALIDVELOCITY_MOVELINABS := 21111,
	NOVALIDACCELERATION_MOVELINABS := 21112,
	NOVALIDDECELERATION_MOVELINABS := 21113,
	NOVALIDJERK_MOVELINABS := 21114,
	TARGETOUTSIDESWLIMITSPASSIVEJOINTS_MOVELINABS := 21115,
	TARGETOUTSIDESWLIMITSMAINAXISX_MOVELINABS := 21116,
	TARGETOUTSIDESWLIMITSMAINAXISY_MOVELINABS := 21117,
	TARGETOUTSIDESWLIMITSMAINAXISZ_MOVELINABS := 21118,
	TARGETOUTSIDESWLIMITSMAINAXISA_MOVELINABS := 21119,
	TARGETOUTSIDESWLIMITSMAINAXISB_MOVELINABS := 21120,
	TARGETOUTSIDESWLIMITSMAINAXISC_MOVELINABS := 21121,
	TARGETOUTSIDESWLIMITSREALAXIS1_MOVELINABS := 21122,
	TARGETOUTSIDESWLIMITSREALAXIS2_MOVELINABS := 21123,
	TARGETOUTSIDESWLIMITSREALAXIS3_MOVELINABS := 21124,
	TARGETOUTSIDESWLIMITSREALAXIS4_MOVELINABS := 21125,
	TARGETOUTSIDESWLIMITSREALAXIS5_MOVELINABS := 21126,
	TARGETOUTSIDESWLIMITSREALAXIS6_MOVELINABS := 21127,
	TARGETOUTSIDESWLIMITSAUXAXIS1_MOVELINABS := 21128,
	TARGETOUTSIDESWLIMITSAUXAXIS2_MOVELINABS := 21129,
	TARGETOUTSIDESWLIMITSAUXAXIS3_MOVELINABS := 21130,
	TARGETOUTSIDESWLIMITSAUXAXIS4_MOVELINABS := 21131,
	TARGETOUTSIDESWLIMITSAUXAXIS5_MOVELINABS := 21132,
	TARGETOUTSIDESWLIMITSAUXAXIS6_MOVELINABS := 21133,
	TARGETTRANSFORMATIONERROR_MOVELINABS := 21134,
	TARGETSINGULARPOS_MOVELINABS := 21135,
	ILLEGALPARAMETER_MOVELINABS := 21136,
	NOVALIDTRANSITIONPARAMETER_MOVELINREL := 21137,
	NOVALIDVELOCITY_MOVELINREL := 21138,
	NOVALIDACCELERATION_MOVELINREL := 21139,
	NOVALIDDECELERATION_MOVELINREL := 21140,
	NOVALIDJERK_MOVELINREL := 21141,
	TARGETOUTSIDESWLIMITSPASSIVEJOINTS_MOVELINREL := 21142,
	TARGETOUTSIDESWLIMITSMAINAXISX_MOVELINREL := 21143,
	TARGETOUTSIDESWLIMITSMAINAXISY_MOVELINREL := 21144,
	TARGETOUTSIDESWLIMITSMAINAXISZ_MOVELINREL := 21145,
	TARGETOUTSIDESWLIMITSMAINAXISA_MOVELINREL := 21146,
	TARGETOUTSIDESWLIMITSMAINAXISB_MOVELINREL := 21147,
	TARGETOUTSIDESWLIMITSMAINAXISC_MOVELINREL := 21148,
	TARGETOUTSIDESWLIMITSREALAXIS1_MOVELINREL := 21149,
	TARGETOUTSIDESWLIMITSREALAXIS2_MOVELINREL := 21150,
	TARGETOUTSIDESWLIMITSREALAXIS3_MOVELINREL := 21151,
	TARGETOUTSIDESWLIMITSREALAXIS4_MOVELINREL := 21152,
	TARGETOUTSIDESWLIMITSREALAXIS5_MOVELINREL := 21153,
	TARGETOUTSIDESWLIMITSREALAXIS6_MOVELINREL := 21154,
	TARGETOUTSIDESWLIMITSAUXAXIS1_MOVELINREL := 21155,
	TARGETOUTSIDESWLIMITSAUXAXIS2_MOVELINREL := 21156,
	TARGETOUTSIDESWLIMITSAUXAXIS3_MOVELINREL := 21157,
	TARGETOUTSIDESWLIMITSAUXAXIS4_MOVELINREL := 21158,
	TARGETOUTSIDESWLIMITSAUXAXIS5_MOVELINREL := 21159,
	TARGETOUTSIDESWLIMITSAUXAXIS6_MOVELINREL := 21160,
	TARGETTRANSFORMATIONERROR_MOVELINREL := 21161,
	TARGETSINGULARPOS_MOVELINREL := 21162,
	ILLEGALPARAMETER_MOVELINREL := 21163,
	NOVALIDTRANSITIONPARAMETER_MOVEDIRABS := 21164,
	DEFAULTVELOCITYOFREALAXISNOTSETMOVEDIRABS := 21165,
	DEFAULTACCELERATIONOFREALAXISNOTSETMOVEDIRABS := 21166,
	DEFAULTDECELERATIONOFREALAXISNOTSETMOVEDIRABS := 21167,
	DEFAULTJERKOFREALAXISNOTSETMOVEDIRABS := 21168,
	TARGETOUTSIDESWLIMITSPASSIVEJOINTS_MOVEDIRABS := 21169,
	TARGETOUTSIDESWLIMITSMAINAXISX_MOVEDIRABS := 21170,
	TARGETOUTSIDESWLIMITSMAINAXISY_MOVEDIRABS := 21171,
	TARGETOUTSIDESWLIMITSMAINAXISZ_MOVEDIRABS := 21172,
	TARGETOUTSIDESWLIMITSMAINAXISA_MOVEDIRABS := 21173,
	TARGETOUTSIDESWLIMITSMAINAXISB_MOVEDIRABS := 21174,
	TARGETOUTSIDESWLIMITSMAINAXISC_MOVEDIRABS := 21175,
	TARGETOUTSIDESWLIMITSREALAXIS1_MOVEDIRABS := 21176,
	TARGETOUTSIDESWLIMITSREALAXIS2_MOVEDIRABS := 21177,
	TARGETOUTSIDESWLIMITSREALAXIS3_MOVEDIRABS := 21178,
	TARGETOUTSIDESWLIMITSREALAXIS4_MOVEDIRABS := 21179,
	TARGETOUTSIDESWLIMITSREALAXIS5_MOVEDIRABS := 21180,
	TARGETOUTSIDESWLIMITSREALAXIS6_MOVEDIRABS := 21181,
	TARGETOUTSIDESWLIMITSAUXAXIS1_MOVEDIRABS := 21182,
	TARGETOUTSIDESWLIMITSAUXAXIS2_MOVEDIRABS := 21183,
	TARGETOUTSIDESWLIMITSAUXAXIS3_MOVEDIRABS := 21184,
	TARGETOUTSIDESWLIMITSAUXAXIS4_MOVEDIRABS := 21185,
	TARGETOUTSIDESWLIMITSAUXAXIS5_MOVEDIRABS := 21186,
	TARGETOUTSIDESWLIMITSAUXAXIS6_MOVEDIRABS := 21187,
	TARGETTRANSFORMATIONERROR_MOVEDIRABS := 21188,
	ILLEGALPARAMETER_MOVEDIRABS := 21189,
	NOVALIDTRANSITIONPARAMETER_MOVEDIRREL := 21190,
	DEFAULTVELOCITYOFREALAXISNOTSETMOVEDIRREL := 21191,
	DEFAULTACCELERATIONOFREALAXISNOTSETMOVEDIRREL := 21192,
	DEFAULTDECELERATIONOFREALAXISNOTSETMOVEDIRREL := 21193,
	DEFAULTJERKOFREALAXISNOTSETMOVEDIRREL := 21194,
	TARGETOUTSIDESWLIMITSPASSIVEJOINTS_MOVEDIRREL := 21195,
	TARGETOUTSIDESWLIMITSMAINAXISX_MOVEDIRREL := 21196,
	TARGETOUTSIDESWLIMITSMAINAXISY_MOVEDIRREL := 21197,
	TARGETOUTSIDESWLIMITSMAINAXISZ_MOVEDIRREL := 21198,
	TARGETOUTSIDESWLIMITSMAINAXISA_MOVEDIRREL := 21199,
	TARGETOUTSIDESWLIMITSMAINAXISB_MOVEDIRREL := 21200,
	TARGETOUTSIDESWLIMITSMAINAXISC_MOVEDIRREL := 21201,
	TARGETOUTSIDESWLIMITSREALAXIS1_MOVEDIRREL := 21202,
	TARGETOUTSIDESWLIMITSREALAXIS2_MOVEDIRREL := 21203,
	TARGETOUTSIDESWLIMITSREALAXIS3_MOVEDIRREL := 21204,
	TARGETOUTSIDESWLIMITSREALAXIS4_MOVEDIRREL := 21205,
	TARGETOUTSIDESWLIMITSREALAXIS5_MOVEDIRREL := 21206,
	TARGETOUTSIDESWLIMITSREALAXIS6_MOVEDIRREL := 21207,
	TARGETOUTSIDESWLIMITSAUXAXIS1_MOVEDIRREL := 21208,
	TARGETOUTSIDESWLIMITSAUXAXIS2_MOVEDIRREL := 21209,
	TARGETOUTSIDESWLIMITSAUXAXIS3_MOVEDIRREL := 21210,
	TARGETOUTSIDESWLIMITSAUXAXIS4_MOVEDIRREL := 21211,
	TARGETOUTSIDESWLIMITSAUXAXIS5_MOVEDIRREL := 21212,
	TARGETOUTSIDESWLIMITSAUXAXIS6_MOVEDIRREL := 21213,
	TARGETTRANSFORMATIONERROR_MOVEDIRREL := 21214,
	ILLEGALPARAMETER_MOVEDIRREL := 21215,
	NOVALIDVELOCITY_MANMODE := 21216,
	NOVALIDACCELERATION_MANMODE := 21217,
	NOVALIDDECELERATION_MANMODE := 21218,
	NOVALIDJERK_MANMODE := 21219,
	MANUALMODEILLEGALPARAMETER := 21220,
	KINEMATICILLEGALPARAMETER := 21221,
	AXESGROUPINERRORSTOP := 21222,
	TOOLINUSE := 21223,
	INVALIDTOOL := 21224,
	AXESGROUPINMOVEMENT := 21225,
	INVALIDCOORDSYSTEM := 21226,
	AXISEXTERNALENABLED := 21227,
	UNSUPPORTEDCOORDSYSTEM := 21228,
	REALAXISNOTREADY := 21229,
	INVALIDAXESGROUPSTATE := 21230,
	REALAXISOUTSIDEWORKINGRANGE := 21231,
	SINGULARPOSITION := 21232,
	L_MC4P_INTERNALERROR := 21233,
	AXESGROUPEXTERNALSTOPPING := 21234,
	RESETAXESGROUPERRORFAILED := 21237,
	ILLEGALTEACHPOSITION := 21238,
	NOTENOUGHMEMORYPATHDATALIST := 21239,
	NOVALIDROTATIONVELOCITY_MOVECIRCABS := 21240,
	NOVALIDROTATIONACCELERATION_MOVECIRCABS := 21241,
	NOVALIDROTATIONJERK_MOVECIRCABS := 21242,
	NOVALIDROTATIONVELOCITY_MOVECIRCREL := 21243,
	NOVALIDROTATIONACCELERATION_MOVECIRCREL := 21244,
	NOVALIDROTATIONJERK_MOVECIRCREL := 21245,
	NOVALIDROTATIONVELOCITY_MOVELINABS := 21246,
	NOVALIDROTATIONACCELERATION_MOVELINABS := 21247,
	NOVALIDROTATIONJERK_MOVELINABS := 21248,
	NOVALIDROTATIONVELOCITY_MOVELINREL := 21249,
	NOVALIDROTATIONACCELERATION_MOVELINREL := 21250,
	NOVALIDROTATIONJERK_MOVELINREL := 21251,
	PATHLIMITVIOLATION_MOVELINABS := 21252,
	PATHLIMITVIOLATION_MOVELINREL := 21253,
	PATHLIMITVIOLATION_MOVECIRCABS := 21254,
	PATHLIMITVIOLATION_MOVECIRCREL := 21255,
	PATHLIMITVIOLATION_MOVEDIRABS := 21256,
	PATHLIMITVIOLATION_MOVEDIRREL := 21257,
	AXESGROUPNOTHOMED := 21258,
	MAINAXISTYPEMODULONOTALLOWED := 21259,
	AXISTYPEMODULONOTALLOWED := 21260,
	AXISLIMITVIOLATIONREALAXIS1VELOCITY := 21261,
	AXISLIMITVIOLATIONREALAXIS2VELOCITY := 21262,
	AXISLIMITVIOLATIONREALAXIS3VELOCITY := 21263,
	AXISLIMITVIOLATIONREALAXIS4VELOCITY := 21264,
	AXISLIMITVIOLATIONREALAXIS5VELOCITY := 21265,
	AXISLIMITVIOLATIONREALAXIS6VELOCITY := 21266,
	AXISLIMITVIOLATIONREALAXIS1ACCELERATION := 21267,
	AXISLIMITVIOLATIONREALAXIS2ACCELERATION := 21268,
	AXISLIMITVIOLATIONREALAXIS3ACCELERATION := 21269,
	AXISLIMITVIOLATIONREALAXIS4ACCELERATION := 21270,
	AXISLIMITVIOLATIONREALAXIS5ACCELERATION := 21271,
	AXISLIMITVIOLATIONREALAXIS6ACCELERATION := 21272,
	AUXAXISSEQUENCEINVALID := 21273,
	AUXAXISNOTALLOWED := 21274,
	ILLEGALTRACKINGPARAMETER := 21275,
	SYNCHRONISATIONERROR := 21276,
	PCSINUSE := 21277,
	TRACKINGFBNOTCALLED := 21278,
	MASTERAXISNOTREADY := 21279,
	MOVEDIRECTNOTALLOWED := 21280,
	AUXAXISNOVALIDVELOCITY := 21281,
	AUXAXISNOVALIDACCELERATION := 21282,
	AUXAXISNOVALIDJERK := 21283,
	MAINAXISNOTCONNECTED := 21284,
	REALAXISNOTCONNECTED := 21285,
	AXESGROUPNOTINITIALIZED := 21286,
	DISABLEDBYPARAMETERTRANSFER := 21287,
	REALAXIS1_ALREADYINUSE := 21288,
	REALAXIS2_ALREADYINUSE := 21289,
	REALAXIS3_ALREADYINUSE := 21290,
	REALAXIS4_ALREADYINUSE := 21291,
	REALAXIS5_ALREADYINUSE := 21292,
	REALAXIS6_ALREADYINUSE := 21293,
	AUXAXIS1_ALREADYINUSE := 21294,
	AUXAXIS2_ALREADYINUSE := 21295,
	AUXAXIS3_ALREADYINUSE := 21296,
	AUXAXIS4_ALREADYINUSE := 21297,
	AUXAXIS5_ALREADYINUSE := 21298,
	AUXAXIS6_ALREADYINUSE := 21299,
	NOVALIDTRANSITIONMODE_MOVECIRCABS := 21300,
	NOVALIDTRANSITIONMODE_MOVECIRCREL := 21301,
	NOVALIDTRANSITIONMODE_MOVELINABS := 21302,
	NOVALIDTRANSITIONMODE_MOVELINREL := 21303,
	NOVALIDTRANSITIONMODE_MOVEDIRABS := 21304,
	NOVALIDTRANSITIONMODE_MOVEDIRREL := 21305,
	NOAXISFORHOMINGSELECTED := 21306,
	INVALIDTARGETORIENTATION := 21307,
	NOKINTRANSFORMATIONAVAILABLE := 21308,
	AXESGROUPNOTSUPPORTED := 21309,
	AXESGROUPNOTDISABLED := 21310,
	AXESGROUPINITFAILED := 21311,
	KINTRANSFORMATIONINUSE := 21312,
	MAXNUMREVOLUTIONSREACHED := 21313,
	PCSCHANGEDDURINGMOTION := 21314,
	CONCURRENTREQUESTMANUALMODE := 21315,
	PATHREFCOMMANDNOTSUPPORTED := 21316,
	PATHREFSYNTAXERROR := 21317,
	PATHREFGCOMMANDNOTSUPPORTED := 21318,
	PATHREFMCOMMANDNOTSUPPORTED := 21319,
	PATHREFINVALIDCOMENTSYNTAX := 21320,
	FILEACCESSTIMEOUT := 21321,
	INVALIDPATHREF := 21322,
	INVALIDPATHFILE := 21323,
	IJKCOMMANDMISSING := 21324,
	INVALIDCIRCCOMMAND := 21325,
	BLENDINGRESETBYINTERNALERROR := 21326,
	DYNAMICCHANGEOFPATHREFNOTALLOWED := 21327,
	CONCURRENTMFUNCTION := 21328,
	INVALIDMFUNCTION := 21329,
	STARTRADIUSGTSEMIMAJORAXIS := 21330,
	STARTRADIUSLTSEMIMINORAXIS := 21331,
	TARGETRADIUSGTSEMIMAJORAXIS := 21332,
	TARGETRADIUSLTSEMIMINORAXIS := 21333,
	SEMIMINORAXISGTSEMIMAJORAXIS := 21334,
	SEMIMINORAXISLE0 := 21335,
	SEMIMAJORAXISLE0 := 21336,
	TARGETNOTONELLIPSE := 21337,
	INVALIDTRAVERSINGRANGECOMBINATION := 21338,
	INVALIDCOORDINATESYSTEMORIENTATION := 21339,
	INVALIDTOOLSYSTEMORIENTATION := 21340,
	TARGETNOTONCIRC := 21341,
	EXECUTIONLOCKEDBYMOVEPATH := 21342,
	NOVALIDVELOCITY_MOVESPLINE := 21343,
	NOVALIDACCELERATION_MOVESPLINE := 21344,
	NOVALIDDECELERATION_MOVESPLINE := 21345,
	NOVALIDJERK_MOVESPLINE := 21346,
	NOVALIDTRANSITIONPARAMETER_MOVESPLINE := 21347,
	NOVALIDTRANSITIONMODE_MOVESPLINE := 21348,
	POSITIONOUTSIDESWLIMITSMAINAXISX_MOVESPLINE := 21349,
	POSITIONOUTSIDESWLIMITSMAINAXISY_MOVESPLINE := 21350,
	POSITIONOUTSIDESWLIMITSMAINAXISZ_MOVESPLINE := 21351,
	POSITIONOUTSIDESWLIMITSMAINAXISA_MOVESPLINE := 21352,
	POSITIONOUTSIDESWLIMITSMAINAXISB_MOVESPLINE := 21353,
	POSITIONOUTSIDESWLIMITSMAINAXISC_MOVESPLINE := 21354,
	NOVALIDROTATIONVELOCITY_MOVESPLINE := 21355,
	NOVALIDROTATIONACCELERATION_MOVESPLINE := 21356,
	NOVALIDROTATIONJERK_MOVESPLINE := 21357,
	NOINTERMEDIATEPOINTS_MOVESPLINE := 21358,
	PATHLIMITVIOLATION_MOVESPLINE := 21359,
	NOVALIDINTERMEDIATEPOINTLOCATION := 21360,
	POSITIONOUTSIDESWLIMITSREALAXIS1_MOVESPLINE := 21361,
	POSITIONOUTSIDESWLIMITSREALAXIS2_MOVESPLINE := 21362,
	POSITIONOUTSIDESWLIMITSREALAXIS3_MOVESPLINE := 21363,
	POSITIONOUTSIDESWLIMITSREALAXIS4_MOVESPLINE := 21364,
	POSITIONOUTSIDESWLIMITSREALAXIS5_MOVESPLINE := 21365,
	POSITIONOUTSIDESWLIMITSREALAXIS6_MOVESPLINE := 21366,
	POSITIONOUTSIDESWLIMITSAUXAXIS1_MOVESPLINE := 21367,
	POSITIONOUTSIDESWLIMITSAUXAXIS2_MOVESPLINE := 21368,
	POSITIONOUTSIDESWLIMITSAUXAXIS3_MOVESPLINE := 21369,
	POSITIONOUTSIDESWLIMITSAUXAXIS4_MOVESPLINE := 21370,
	POSITIONOUTSIDESWLIMITSAUXAXIS5_MOVESPLINE := 21371,
	POSITIONOUTSIDESWLIMITSAUXAXIS6_MOVESPLINE := 21372,
	POSITIONTRANSFORMATIONERROR_MOVESPLINE := 21373,
	POSITIONOUTSIDESWLIMITSPASSIVEJOINTS_MOVESPLINE := 21374,
	POSITIONSINGULARPOS_MOVESPLINE := 21375,
	CONCURRENTTORQUEPRECONTROL := 21376,
	INVALIDORIENTATIONMODE := 21377,
	CONCURRENTAXESGROUPBASICCONTROL := 21378,
	PARAMETERLIMITSNOTSUFFICIENT := 21379,
	SETVALUEMANIPULATIONNOTSUPPORTED := 21380,
	MINPOSGTMAXPOS := 21381,
	DYNAMICPARAMETERNOTPLAUSIBLE := 21382,
	CONVERGENCENOTSUFFICIENT := 21383,
	IDENTIFICATIONNOTDONE := 21384,
	INVALIDOVERRIDEFORIDENTIFICATION := 21385,
	DUALUSELICENSEMISSING := 21386,
	CONCURRENTMOVEPATH := 21387,
	MAINAXISNOTSUPPORTED := 21389,
	BLENDINGCARTESIANWITHMOVEDIRECTNOTSUPPORTED := 21390,
	BLENDINGWAITTIMENOTSUPPORTED := 21391,
	BLENDINGAUXILLIARYAXESNOTSUPPORTED := 21392,
	BLENDINGRESETNOPREDECESSOR := 21393,
	BLENDINGRESETEXECUTETOOLATE := 21394,
	BLENDINGRESETLOOKAHEADZERO := 21395,
	PATHREFABORTED := 21396,
	BLENDINGRESETTOOLCHANGED := 21397,
	INVALIDSWITCHTIME := 21398,
	INVALIDGOTOTARGET := 21399,
	RECURSIVESUBROUTINECALL := 21400,
	SUBROUTINEDEPTHEXCEEDED := 21401,
	INVALIDSUBROUTINESYNTAX := 21402,
	INVALIDMFUNTYPEFORINTERPRETERHALT := 21403,
	FINISHDATAINCONSISTENT := 21404,
	FINISHNOTPOSSIBLEABORTDURINGPATHPREP := 21405,
	CMDSYNCINSTARTREQUIRED := 21406,
	INVALIDTRACKINGOBJECT := 21407,
	CONCURRENTCMDSYNCINSTART := 21408,
	INVALIDCOORDSYSTEMFORTRACKING := 21409,
	MOVECMDFORTRACKINGREQUIRED := 21410,
	CONCURRENTDIGITALSWITCHHANDLER := 21411,
	NOPARAMFORHFUN := 21412,
	MOVECMDREQUIREDFORHFUN := 21413,
	OPARAMREQUIREDFORG00WITHHFUN := 21414,
	OPARAMREQUIREDFORG04WITHHFUN := 21415,
	CONCURRENTPARAMFORHFUN := 21416,
	HFUNREQIREDFORLPARAM := 21417,
	HFUNREQIREDFOROPARAM := 21418,
	HFUNVALUEOUTOFRANGE := 21419,
	NUMBEROFALLOWEDHFUNEXCEEDED := 21420,
	CONCURRENTREGULATORON := 21421,
	CONCURRENTENABLEOPERATION := 21422,
	PATHVELOCITYLIMITED := 21423,
	PATHACCELERATIONLIMITED := 21424,
	PATHJERKLIMITED := 21425,
	PHASINGNOTALLOWED := 22000,
	INVALIDCAMREF := 22010,
	INVALIDCAMTYPE := 22011,
	INVALIDCAMDATA := 22012,
	INVALIDDATACOUNT := 22013,
	DATACOUNTTOOSMALL := 22014,
	INVALIDLAWOFMOTION := 22015,
	INVALIDINPUTDATA := 22016,
	MASTEROUTOFCAM := 22025,
	INVALIDVELACC_OFFSETSCALING := 22026,
	INVALIDCAMTABLE := 22027,
	INVALIDSTARTORENDPOSOFCAM := 22028,
	INVALIDSCALINGFACTOR := 22029,
	RAMPINERROR := 22030,
	NOTALLOWEDMOVEMENTBYMASTER := 22035,
	CLUTCHISREVERSING := 22036,
	INVALIDDEFAULTJERK := 22037,
	INVALIDOPENINSTANTDEC := 22038,
	INVALIDREVERSE := 22039,
	FILENOTFOUND := 22050,
	INVALIDFILE := 22051,
	INVALIDCHECKCRC := 22052,
	INVALIDDATASIZE := 22053,
	INVALIDTAPPETREF := 22060,
	INVALIDTAPPETDATA := 22061,
	INVALIDTAPPETTYPE := 22062,
	INVALIDTIMINGTAPPET := 22063,
	INVALIDPOSSELECTIONTAPPET := 22064,
	DYNAMISATIONERROR := 22065,
	XCYCLELENGTHINVALID_LINEARCOUPLING := 22082,
	YCYCLELENGTHINVALID_LINEARCOUPLING := 22083,
	POSININVALID_LINEARCOUPLING := 22084,
	INVALIDTAPPETSCOUNT := 22085,
	RESETPHASINGNOTALLOWED := 22086,
	INVALIDMASTERSYNCPOSITION := 22087,
	INVALIDSCALINGOFFSETMODE := 22089,
	INVALIDCOMBINEMODE := 22090,
	INVALIDSYNCMODE := 22091,
	INVALIDERRORHANDLER := 23001,
	INVALIDERRORID := 23002,
	INVALIDTEXTREFID := 23003,
	INVALIDDEFAULTTEXTREFID := 23004,
	INVALIDPOINTERERRORMSGBUFFER := 23050,
	INVALIDBUFFERSIZEERRORMSGBUFFER := 23051,
	INVALIDSTARTORENDINDEX := 23052,
	ERRMSGBUFFERDATATOOSMALL := 23053,
	ERRORMSGLISTNOTAVAILABLE := 23054,
	ERRORMSGLISTNOTACCESSIBLE := 23055,
	NUMBERSUPPORTPOINTSEXCEEDED := 24001,
	STRICLYMONOTONINCREASINGVALUESREQUIRED := 24002,
	INVALIDARRAYBOUND := 24003,
	ARRAYBOUNDSMISMATCH := 24004,
	SINGULARMATRIX := 24005,
	INVALIDINTERPOLATIONTYPE := 24006,
	SYSLOGNOTAVAILABLE := 25001,
	NOSYSLOGRESOURCEAVAILABLE := 25002,
	SYSLOGINVALIDSPECIALCHARACTER := 25003,
	FUNCTIONMODULENOTCONNECTED := 26001,
	DEVICEMODULENOTCONNECTED := 26002,
	FUNCTIONMODULENOTSUPPORTED := 26003,
	DEVICEMODULENOTSUPPORTED := 26004,
	NOTSUPPORTEDBYMODULEHANDLERVERSION := 26005,
	INVALIDDISCONNECTMODE := 26006,
	DEVICEALREADYCONNECTED := 26007,
	AXISCALLNOTINMOTIONTASK := 26501,
	POUCALLNOTINMOTIONTASK := 26502,
	POUCALLTWICE := 26503,
	POUCALLMORETHANTWICE := 26504,
	TASKASSIGNMENTMISMATCH := 26505,
	SKEWNESSMONITORINGWARNING := 27000,
	SKEWNESSMONITORINGERROR := 27001,
	TENSIONMONITORINGWARNING := 27002,
	TENSIONMONITORINGERROR := 27003,
	MAINAXISALREADYASSIGNED := 27004,
	FOLLOWINGAXISALREADYASSIGNED := 27005,
	SELECTEDAXISALREADYINUSE := 27006,
	NOTREADYFORALIGNMENT := 27008,
	MAINAXISINERROR := 27009,
	FOLLOWINGAXISINERROR := 27010,
	KINEMATICINERROR := 27011,
	NOAXISSELECTED := 27012,
	FOLLOWINGAXISNOTSELECTED := 27013,
	MAINAXISNOTSELECTED := 27014,
	MAINANDFOLLOWINGAXISIDENTICAL := 27015,
	FOLLOWINGAXISALREADYUSED := 27016,
	FUNCTIONNOTSUPPORTEDFORFOLLOWINGAXIS := 27017,
	AXISCONFIGNOTEQUALHOMINGMODE := 27019,
	INVALIDHOMINGSEQUENCE := 27020,
	DIFFERENTHOMINGPARAMETER := 27021,
	FUNCTIONNOTSUPPORTEDBYCONTROLLERFW := 28000,
	COMPONENTNAMENOTFOUND := 28001,
	ETHERCATMASTERNOTAVAILABLE := 28500
);
END_TYPE

(* ---- L_IE1P_ERRORDATA.dut ---- *)
TYPE L_IE1P_ERRORDATA :
STRUCT
	INSTANCEID : UDINT;
	TEXTREFID : UINT;
	EVENTID : UINT;
	SEVERITY : USINT;
	LAYER : USINT;
	STATE : USINT;
	DUMMY : USINT;
END_STRUCT
END_TYPE

(* ---- L_IE1P_GROUP.dut ---- *)
TYPE L_IE1P_GROUP :
(
	USERGROUP1 := 1,
	USERGROUP2 := 2,
	USERGROUP3 := 3,
	USERGROUP4 := 4,
	USERGROUP5 := 5,
	MANUFACTURERGROUP := 12
);
END_TYPE

(* ---- L_IE1P_REACTION.dut ---- *)
TYPE L_IE1P_REACTION :
(
	NO_REACTION := 0,
	USERREACTION1 := 1,
	USERREACTION2 := 2,
	CYCLESTOP := 3,
	NORMALSTOP := 4,
	FASTSTOP := 5,
	USERREACTION6 := 6,
	QSPAPPL := 11,
	QSP := 12,
	QSP_CINH := 13,
	CINH := 14
);
END_TYPE

(* ---- L_IE1P_REACTIONCOUNTER.dut ---- *)
TYPE L_IE1P_REACTIONCOUNTER :
STRUCT
	USERREACTION1 : DINT;
	USERREACTION2 : DINT;
	CYCLESTOP : DINT;
	NORMALSTOP : DINT;
	FASTSTOP : DINT;
	USERREACTION6 : DINT;
	QSPAPPL : DINT;
	QSP : DINT;
	QSP_CINH : DINT;
	CINH : DINT;
END_STRUCT
END_TYPE

(* ---- L_IE1P_REACTIONSTATUS.dut ---- *)
TYPE L_IE1P_REACTIONSTATUS :
STRUCT
	USERREACTION1 : BOOL;
	USERREACTION2 : BOOL;
	CYCLESTOP : BOOL;
	NORMALSTOP : BOOL;
	FASTSTOP : BOOL;
	USERREACTION6 : BOOL;
	QSPAPPL : BOOL;
	QSP : BOOL;
	QSP_CINH : BOOL;
	CINH : BOOL;
END_STRUCT
END_TYPE

(* ---- L_IE1P_READERRORDATA.dut ---- *)
TYPE L_IE1P_READERRORDATA :
STRUCT
	NUMBEROFENTRIES : DWORD;
	CMPERRORDATA : ARRAY [1..1000] OF L_IE1P_ErrorData;
END_STRUCT
END_TYPE

(* ---- L_IE1P_SERVERITYLEVEL.dut ---- *)
TYPE L_IE1P_SERVERITYLEVEL :
(
	NO_RESPONSE := 0,
	WARNING := 2,
	INFORMATION := 11,
	WARNING_LOCK := 13,
	FAULT_QSPAPPL := 19,
	FAULT_QSP := 20,
	FAULT_QSP_CINH := 21,
	FAULT := 23
);
END_TYPE

(* ---- L_IE1P_SEVERITYCOUNTER.dut ---- *)
TYPE L_IE1P_SEVERITYCOUNTER :
STRUCT
	WARNING : DINT;
	INFORMATION : DINT;
	WARNING_LOCK : DINT;
	FAULT_LOG : DINT;
	FAULT_QSPAPPL : DINT;
	FAULT_QSP : DINT;
	FAULT_QSP_CINH : DINT;
	FAULT_CINH : DINT;
	FAULT : DINT;
END_STRUCT
END_TYPE

(* ---- L_IE1P_SEVERITYLEVEL.dut ---- *)
TYPE L_IE1P_SEVERITYLEVEL :
(
	NO_RESPONSE := 0,
	WARNING := 2,
	INFORMATION := 11,
	WARNING_LOCK := 13,
	FAULT_LOG := 18,
	FAULT_QSPAPPL := 19,
	FAULT_QSP := 20,
	FAULT_QSP_CINH := 21,
	FAULT_CINH := 23,
	FAULT := 30
);
END_TYPE

(* ---- L_IE1P_SEVERITYSTATUS.dut ---- *)
TYPE L_IE1P_SEVERITYSTATUS :
STRUCT
	WARNING : BOOL;
	INFORMATION : BOOL;
	WARNING_LOCK : BOOL;
	FAULT_LOG : BOOL;
	FAULT_QSPAPPL : BOOL;
	FAULT_QSP : BOOL;
	FAULT_QSP_CINH : BOOL;
	FAULT_CINH : BOOL;
	FAULT : BOOL;
END_STRUCT
END_TYPE

(* ---- GVL.gvl ---- *)
VAR_GLOBAL
END_VAR

(* ---- L_IE1P_IERRORHANDLER.itf ---- *)
INTERFACE L_IE1P_IERRORHANDLER
END_INTERFACE

METHOD ITFCHECKERRORRESETOCCURED : BOOL
VAR_IN_OUT
	RESETTIME : SYSTIME;
END_VAR
END_METHOD

METHOD ITFCLEARERROR : DWORD
VAR_INPUT
	ESEVERITY : L_IE1P_SeverityLevel;
	WERRORID : WORD;
	WCOMPID : WORD;
	DWINSTANCEID : DWORD := 0;
END_VAR
END_METHOD

METHOD ITFCLEARREACTION
VAR_INPUT
	EREACTION : L_IE1P_Reaction;
	DICLEARCOUNT : DINT;
	DWINSTANCEID : DWORD;
END_VAR
END_METHOD

METHOD ITFGETACTUALERRORCODE : DWORD
VAR_OUTPUT
	ESEVERITY : WORD;
END_VAR
END_METHOD

METHOD ITFREGISTERERRORINSTANCE : DWORD
END_METHOD

METHOD ITFRESETACTIVE : BOOL
END_METHOD

METHOD ITFRESETERROR : DWORD
VAR_INPUT
	ERRORHANDLE : RTS_IEC_HANDLE := 0;
END_VAR
END_METHOD

METHOD ITFRESETERRORREACTION
VAR_INPUT
	DWINSTANCEID : DWORD := 0;
END_VAR
END_METHOD

METHOD ITFSETERROR : DWORD
VAR_INPUT
	ESEVERITY : L_IE1P_SeverityLevel;
	WERRORID : WORD;
	WCOMPID : WORD;
	DWINSTANCEID : DWORD := 0;
	EREACTION : L_IE1P_Reaction;
END_VAR
END_METHOD

(* ---- GETBOOLEANPROPERTY.pou ---- *)
FUNCTION GETBOOLEANPROPERTY : BOOL
VAR_INPUT
	STKEY : WSTRING;
END_VAR
END_FUNCTION

(* ---- GETCOMPANY.pou ---- *)
FUNCTION GETCOMPANY : WSTRING
END_FUNCTION

(* ---- GETNUMBERPROPERTY.pou ---- *)
FUNCTION GETNUMBERPROPERTY : DINT
VAR_INPUT
	STKEY : WSTRING;
END_VAR
END_FUNCTION

(* ---- GETTEXTPROPERTY.pou ---- *)
FUNCTION GETTEXTPROPERTY : WSTRING
VAR_INPUT
	STKEY : WSTRING;
END_VAR
END_FUNCTION

(* ---- GETTEXTPROPERTY2.pou ---- *)
FUNCTION GETTEXTPROPERTY2 : POINTER TO WSTRING
VAR_INPUT
	STKEY : WSTRING;
END_VAR
END_FUNCTION

(* ---- GETTITLE.pou ---- *)
FUNCTION GETTITLE : WSTRING
END_FUNCTION

(* ---- GETVERSION.pou ---- *)
FUNCTION GETVERSION : VERSION
END_FUNCTION

(* ---- GETVERSIONPROPERTY.pou ---- *)
FUNCTION GETVERSIONPROPERTY : VERSION
VAR_INPUT
	STKEY : WSTRING;
END_VAR
END_FUNCTION

(* ---- LENZEERRMGR_11264.pou ---- *)
FUNCTION_BLOCK LENZEERRMGR_11264
VAR
	M_TEXTLISTFILE : STRING(255);
	_STNAMESPACE : STRING;
END_VAR
END_FUNCTION_BLOCK
